(* PLC project , Example Fixture *)

FUNCTION_BLOCK FB_Cmd
  VAR_INPUT
    Cmd : BOOL;
    Ack : BOOL;
  END_VAR
  VAR_OUTPUT
    Busy : BOOL;
  END_VAR

(* LD diagram, written out as Structured Text *)
Cmd := Ack;
Busy := Cmd;
END_FUNCTION_BLOCK

CONFIGURATION c
  RESOURCE r ON PLC
  END_RESOURCE
END_CONFIGURATION
